Yaskawa INFORM job: -DEFRO-70-PRZYLACZE-70KASUJ.JBI

/JOB
//NAME -DEFRO-70-PRZYLACZE-70KASUJ
//POS
///NPOS 124,124,124,0,0,0
///TOOL 0
///POSTYPE PULSE
///PULSE
C00000=-283,-101162,-84213,3710,-80188,-1936
C00001=-283,-101162,-84213,3710,-80188,-1936
C00002=116617,-39062,-41553,1138,-40446,20
C00003=129312,23670,-33720,-14256,-61435,76595
C00004=149817,31841,-31795,27011,-57385,28137
C00005=152773,60456,-9717,30826,-76450,24874
C00006=149980,46799,-17890,30362,-63313,13597
C00007=141160,51169,-7378,14366,-65778,3091
C00008=136677,64016,6397,6150,-76179,-494
C00009=141378,9053,-49023,24268,-47565,-67133
C00010=125496,48327,-10508,-10752,-65084,-13725
C00011=130369,56785,-528,-1011,-71593,-13969
C00012=129107,53038,-4370,-2924,-69346,-18638
C00013=128986,13733,-25067,-13195,-71631,75488
C00014=115254,13128,-25616,-11802,-73565,79847
C00015=115259,22487,-34865,-12640,-63289,80918
C00016=131340,5225,-55572,19882,-37557,40272
C00017=141113,50251,-21422,35156,-71250,27064
C00018=141007,50182,-21498,35193,-71206,27085
C00019=141007,50182,-21498,35193,-71206,27085
C00020=137714,37646,-27763,32896,-58429,16473
C00021=129076,45247,-14016,15951,-62855,6645
C00022=121365,54735,-2868,3704,-70570,-4230
C00023=105889,56250,-7649,-21324,-75365,-25403
C00024=98023,31978,-40039,-45182,-56261,-13451
C00025=100224,44212,-25129,-32797,-73818,-42058
C00026=102299,40629,-26008,-28475,-71942,-45909
C00027=121076,21343,-35316,908,-62246,-81562
C00028=121076,10747,-22159,833,-75786,-81463
C00029=100383,18918,-18562,-9881,-76761,84439
C00030=101335,27463,-29788,-10664,-65529,85098
C00031=115713,4222,-56662,15198,-34727,46918
C00032=128373,44829,-27529,39504,-66240,29595
C00033=124328,33310,-32072,34883,-53820,19937
C00034=124328,33310,-32072,34883,-53820,19937
C00035=116075,45486,-13239,16661,-61560,10020
C00036=112317,60890,2820,11495,-73723,-606
C00037=94613,64601,2142,-17801,-79259,-22601
C00038=91137,54103,-11116,-25365,-70739,-18946
C00039=86945,42270,-27280,-36642,-61219,-13206
C00040=88301,54680,-13566,-28329,-78742,-39649
C00041=93612,48687,-14019,-16896,-75888,-44120
C00042=107037,24185,-32573,2312,-62235,-77114
C00043=100383,18918,-18562,-9881,-76761,84439
C00044=88082,30336,-7531,-8088,-78954,88284
C00045=89154,35127,-22112,-8522,-65087,85240
C00046=89544,34712,-22538,-8576,-65002,85121
C00047=100203,10236,-51959,9142,-32676,54086
C00048=115214,43849,-28542,43438,-61422,32379
C00049=110430,34623,-30597,35948,-49426,23884
C00050=101177,66932,10039,13677,-73518,2856
C00051=84754,73517,14044,-12253,-80824,-22539
C00052=78238,80066,13225,-23326,-87649,-28956
C00053=78238,80066,13225,-23326,-87649,-28956
C00054=77744,70007,4024,-24183,-84112,-37607
C00055=93905,32013,-24678,3546,-62668,-72921
C00056=93951,24843,-16667,3331,-71267,-72683
C00057=77831,45702,7684,-6459,-81284,91476
C00058=78073,52891,-3303,-6771,-70880,91958
C00059=86321,21390,-41402,2747,-32621,60915
C00060=102328,48592,-23384,46468,-56980,35399
C00061=97622,41313,-23800,35801,-45769,27976
C00062=95336,65754,6791,24352,-65412,15878
C00063=90551,78368,23842,15429,-74357,6364
C00064=75321,97136,42564,-11419,-90206,-17945
C00065=66680,76750,12803,-30175,-73528,-10031
C00066=68858,90162,29080,-20673,-90872,-36103
C00067=68858,90162,29080,-20673,-90872,-36103
C00068=68890,88039,27277,-20264,-89888,-36525
C00069=82457,45121,-10983,4500,-63864,-69204
C00070=77831,46763,5255,-6493,-79257,91580
C00071=100383,18918,-18562,-9881,-76761,84439
C00072=124101,-43184,-98243,-16518,52281,7000
C00073=123755,-7958,-89511,-14194,64535,5137
C00074=123755,-7958,-89511,-14194,64535,5137
C00075=120912,-12617,-93089,-9839,60859,10956
C00076=121533,-31212,-92910,-11510,35078,6544
C00077=122206,-29072,-90087,-12243,35589,-2657
C00078=123755,-7840,-89515,-14187,64596,5129
C00079=123755,-27930,-86554,-16069,52849,6788
C00080=123755,-31596,-85257,-16659,50271,7220
C00081=123755,-28371,-86416,-16134,52549,6837
C00082=123755,-7958,-89511,-14194,64535,5137
C00083=121932,-4467,-89644,-7852,68214,10996
C00084=130594,-5675,-87742,-32640,65606,16968
C00085=121207,-33956,-80021,-42944,8634,21416
C00086=121398,-33051,-89073,-12931,27077,-1891
C00087=119830,-29976,-89766,-6946,33011,-10480
C00088=121383,9671,-86957,-7975,82780,3273
C00089=123844,-33214,-84175,-16864,48398,7942
C00090=123999,-39711,-94755,-16482,51917,7023
C00091=123520,-8018,-89739,-13952,64610,5074
C00092=123514,-7754,-89533,-13967,64621,5071
C00093=125747,-8511,-91196,-20044,64124,16767
C00094=124758,-33497,-85798,-35788,21508,19109
C00095=121444,-34263,-87472,-15236,22128,1720
C00096=117635,-29901,-89670,2040,32900,-12364
C00097=120806,-19229,-91385,-7013,51591,-4269
C00098=123278,-3298,-89359,-12226,69976,6390
C00099=123735,-32674,-90978,-15994,53118,6740
C00100=123835,-44294,-91959,-17334,47983,7666
C00101=122869,-6543,-89983,-11258,66473,7782
C00102=122869,-6622,-89981,-11262,66432,7786
C00103=120666,-24161,-92251,-9656,44301,18332
C00104=120622,-35099,-88572,-13686,22135,5149
C00105=121670,-32826,-90694,-12460,29863,-58
C00106=120799,-29821,-90097,-9101,34108,-7769
C00107=117992,-25289,-89559,-1030,40191,-9143
C00108=122619,-6933,-90139,-10800,66466,8097
C00109=122622,-7156,-90314,-10803,66459,8098
C00110=123632,-25499,-87776,-15569,54758,6451
C00111=123637,-32760,-85682,-16630,49927,7238
C00112=123766,-34030,-92143,-16017,53144,6747
C00113=122032,-5500,-90078,-8484,67787,10331
C00114=122032,-5500,-90078,-8484,67787,10331
C00115=119888,-26436,-91823,-7086,40086,20761
C00116=120072,-35228,-83770,-17836,12895,7656
C00117=119245,-35145,-84473,-5873,14566,-1771
C00118=120774,-28613,-91055,-8481,37254,-8445
C00119=122137,-20625,-91389,-11840,49625,-8457
C00120=122281,3827,-88512,-9548,77692,7214
C00121=124756,-84422,-108366,-22045,38231,10349
C00122=2454,-100942,-83171,2490,-79441,1084
C00123=-283,-101162,-84213,3710,-80188,-1936
BC00000=570125
BC00001=954451
BC00002=878037
BC00003=914864
BC00004=914864
BC00005=914864
BC00006=914864
BC00007=914864
BC00008=914864
BC00009=914864
BC00010=914864
BC00011=914864
BC00012=914864
BC00013=914864
BC00014=914864
BC00015=914864
BC00016=914864
BC00017=914864
BC00018=914864
BC00019=914864
BC00020=914864
BC00021=914864
BC00022=914864
BC00023=914864
BC00024=914864
BC00025=914864
BC00026=914864
BC00027=914864
BC00028=914864
BC00029=914864
BC00030=914864
BC00031=914864
BC00032=914864
BC00033=914864
BC00034=914864
BC00035=914864
BC00036=914864
BC00037=914863
BC00038=914863
BC00039=914864
BC00040=914864
BC00041=914864
BC00042=914864
BC00043=914864
BC00044=914864
BC00045=914864
BC00046=914864
BC00047=914864
BC00048=914864
BC00049=914864
BC00050=914864
BC00051=914864
BC00052=914864
BC00053=914864
BC00054=914864
BC00055=914864
BC00056=914864
BC00057=914864
BC00058=914864
BC00059=914864
BC00060=914864
BC00061=914864
BC00062=914864
BC00063=914864
BC00064=914863
BC00065=914864
BC00066=914864
BC00067=914864
BC00068=914864
BC00069=914864
BC00070=914864
BC00071=914864
BC00072=869720
BC00073=869720
BC00074=869720
BC00075=869720
BC00076=869720
BC00077=869720
BC00078=869720
BC00079=869720
BC00080=869720
BC00081=908129
BC00082=908129
BC00083=908129
BC00084=907961
BC00085=908580
BC00086=908293
BC00087=908102
BC00088=907757
BC00089=908179
BC00090=945847
BC00091=945846
BC00092=945847
BC00093=946325
BC00094=946857
BC00095=946662
BC00096=946390
BC00097=946210
BC00098=945983
BC00099=945983
BC00100=984509
BC00101=984509
BC00102=984509
BC00103=984689
BC00104=985047
BC00105=984920
BC00106=984769
BC00107=984449
BC00108=984290
BC00109=984290
BC00110=984290
BC00111=1022837
BC00112=1022864
BC00113=1022864
BC00114=1022864
BC00115=1022915
BC00116=1023549
BC00117=1023332
BC00118=1022983
BC00119=1022931
BC00120=1022837
BC00121=1022837
BC00122=1040800
BC00123=570125
EC00000=1166,0
EC00001=1166,0
EC00002=-1743,0
EC00003=-1741,0
EC00004=-1741,0
EC00005=-1741,0
EC00006=-1740,0
EC00007=-1740,0
EC00008=-1740,0
EC00009=-1740,0
EC00010=-1740,0
EC00011=-1740,0
EC00012=-1740,0
EC00013=-1741,0
EC00014=-1741,0
EC00015=-1741,0
EC00016=-1741,0
EC00017=-1741,0
EC00018=-1741,0
EC00019=-1741,0
EC00020=-1740,0
EC00021=-1740,0
EC00022=-1740,0
EC00023=-1740,0
EC00024=-1740,0
EC00025=-1741,0
EC00026=-1741,0
EC00027=-1740,0
EC00028=-1740,0
EC00029=-1741,0
EC00030=-1741,0
EC00031=-1741,0
EC00032=-1741,0
EC00033=-1741,0
EC00034=-1741,0
EC00035=-1740,0
EC00036=-1740,0
EC00037=-1741,0
EC00038=-1741,0
EC00039=-1740,0
EC00040=-1741,0
EC00041=-1741,0
EC00042=-1740,0
EC00043=-1741,0
EC00044=-1741,0
EC00045=-1741,0
EC00046=-1741,0
EC00047=-1741,0
EC00048=-1741,0
EC00049=-1741,0
EC00050=-1740,0
EC00051=-1741,0
EC00052=-1741,0
EC00053=-1741,0
EC00054=-1741,0
EC00055=-1740,0
EC00056=-1740,0
EC00057=-1741,0
EC00058=-1741,0
EC00059=-1741,0
EC00060=-1741,0
EC00061=-1741,0
EC00062=-1740,0
EC00063=-1740,0
EC00064=-1741,0
EC00065=-1740,0
EC00066=-1741,0
EC00067=-1741,0
EC00068=-1741,0
EC00069=-1740,0
EC00070=-1741,0
EC00071=-1741,0
EC00072=-85617,0
EC00073=-85617,0
EC00074=-85617,0
EC00075=-85617,0
EC00076=-85617,0
EC00077=-85617,0
EC00078=-85617,0
EC00079=-85617,0
EC00080=-85617,0
EC00081=-85617,0
EC00082=-85617,0
EC00083=-85617,0
EC00084=-85617,0
EC00085=-85617,0
EC00086=-85617,0
EC00087=-85617,0
EC00088=-85617,0
EC00089=-85617,0
EC00090=-85617,0
EC00091=-85617,0
EC00092=-85617,0
EC00093=-85617,0
EC00094=-85617,0
EC00095=-85617,0
EC00096=-85617,0
EC00097=-85617,0
EC00098=-85617,0
EC00099=-85617,0
EC00100=-85617,0
EC00101=-85617,0
EC00102=-85617,0
EC00103=-85617,0
EC00104=-85617,0
EC00105=-85617,0
EC00106=-85617,0
EC00107=-85617,0
EC00108=-85617,0
EC00109=-85617,0
EC00110=-85617,0
EC00111=-85617,0
EC00112=-85617,0
EC00113=-85617,0
EC00114=-85617,0
EC00115=-85617,0
EC00116=-85617,0
EC00117=-85617,0
EC00118=-85617,0
EC00119=-85617,0
EC00120=-85617,0
EC00121=-85617,0
EC00122=946,0
EC00123=1166,0
//INST
///DATE 2025/05/08 13:43
///COMM OZZ
///ATTR SC,RW
///GROUP1 RB1,BS1
///GROUP2 ST1
NOP
MOVJ C00000 BC00000 VJ=70.00 DEC=20  +MOVJ EC00000 VJ=70.00
MOVJ C00001 BC00001 VJ=40.00 DEC=20  +MOVJ EC00001 VJ=40.00
MOVJ C00002 BC00002 VJ=70.00 DEC=20  +MOVJ EC00002 VJ=70.00
MOVJ C00003 BC00003 VJ=80.00 DEC=20  +MOVJ EC00003 VJ=80.00
MACRO1 MJ#(0) ARGF10
WVON WEV#(2)
ARCON
MOVL C00004 BC00004 V=5.0 DEC=20  +MOVJ EC00004 VJ=80.00
MOVC C00005 BC00005 V=5.0 DEC=20  +MOVJ EC00005 VJ=80.00
WVON WEV#(1)
MOVC C00006 BC00006 V=5.0 DEC=20  +MOVJ EC00006 VJ=80.00
MOVC C00007 BC00007 V=5.0 DEC=20  +MOVJ EC00007 VJ=80.00
MOVC C00008 BC00008 V=5.0 DEC=20  +MOVJ EC00008 VJ=80.00
MOVC C00009 BC00009 V=5.0 DEC=20  +MOVJ EC00009 VJ=80.00
MOVL C00010 BC00010 V=5.0 DEC=20  +MOVJ EC00010 VJ=80.00
MOVC C00011 BC00011 V=5.0 DEC=20  +MOVJ EC00011 VJ=80.00
MOVL C00012 BC00012 V=5.0 DEC=20  +MOVJ EC00012 VJ=80.00
WVOF
ARCOF
MOVJ C00013 BC00013 VJ=80.00 DEC=20  +MOVJ EC00013 VJ=80.00
MOVJ C00014 BC00014 VJ=80.00 DEC=20  +MOVJ EC00014 VJ=80.00
MOVJ C00015 BC00015 VJ=80.00 DEC=20  +MOVJ EC00015 VJ=0.78
MACRO1 MJ#(0) ARGF10
WVON WEV#(2)
ARCON
MOVC C00016 BC00016 V=5.0 DEC=20  +MOVJ EC00016 VJ=40.00
MOVL C00017 BC00017 V=5.0 DEC=20  +MOVJ EC00017 VJ=40.00
WVON WEV#(1)
MOVC C00018 BC00018 V=1500.0 DEC=20  +MOVJ EC00018 VJ=40.00
MOVC C00019 BC00019 V=600.0 DEC=20  +MOVJ EC00019 VJ=40.00
MOVC C00020 BC00020 V=5.0 DEC=20  +MOVJ EC00020 VJ=40.00
MOVC C00021 BC00021 V=5.0 DEC=20  +MOVJ EC00021 VJ=100.00
MOVC C00022 BC00022 V=5.0 DEC=20  +MOVJ EC00022 VJ=40.00
MOVC C00023 BC00023 V=5.0 DEC=20  +MOVJ EC00023 VJ=40.00
MOVL C00024 BC00024 V=5.0 DEC=20  +MOVJ EC00024 VJ=40.00
WVON WEV#(2)
MOVC C00025 BC00025 V=5.0 DEC=20  +MOVJ EC00025 VJ=40.00
MOVC C00026 BC00026 V=5.0 DEC=20  +MOVJ EC00026 VJ=80.00
MOVC C00027 BC00027 V=5.0 DEC=20  +MOVJ EC00027 VJ=40.00
WVOF
ARCOF
MOVJ C00028 BC00028 VJ=80.00 DEC=20  +MOVJ EC00028 VJ=80.00
MOVJ C00029 BC00029 VJ=80.00 DEC=20  +MOVJ EC00029 VJ=80.00
MOVJ C00030 BC00030 VJ=80.00 DEC=20  +MOVJ EC00030 VJ=80.00
MACRO1 MJ#(0) ARGF10
WVON WEV#(2)
ARCON
MOVC C00031 BC00031 V=5.0 DEC=20  +MOVJ EC00031 VJ=80.00
MOVL C00032 BC00032 V=5.0 DEC=20  +MOVJ EC00032 VJ=80.00
WVON WEV#(1)
MOVC C00033 BC00033 V=5.0 DEC=20  +MOVJ EC00033 VJ=80.00
MOVL C00034 BC00034 V=5.0 DEC=20  +MOVJ EC00034 VJ=80.00
MOVC C00035 BC00035 V=5.0 DEC=20  +MOVJ EC00035 VJ=80.00
MOVC C00036 BC00036 V=5.0 DEC=20  +MOVJ EC00036 VJ=80.00
MOVC C00037 BC00037 V=5.0 DEC=20  +MOVJ EC00037 VJ=80.00
MOVC C00038 BC00038 V=5.0 DEC=20  +MOVJ EC00038 VJ=80.00
MOVL C00039 BC00039 V=5.0 DEC=20  +MOVJ EC00039 VJ=80.00
MOVC C00040 BC00040 V=5.0 DEC=20  +MOVJ EC00040 VJ=80.00
MOVC C00041 BC00041 V=5.0 DEC=20  +MOVJ EC00041 VJ=80.00
MOVC C00042 BC00042 V=5.0 DEC=20  +MOVJ EC00042 VJ=80.00
WVOF
ARCOF
MOVJ C00043 BC00043 VJ=80.00 DEC=20  +MOVJ EC00043 VJ=80.00
MOVJ C00044 BC00044 VJ=80.00 DEC=20  +MOVJ EC00044 VJ=80.00
MOVJ C00045 BC00045 VJ=80.00 DEC=20  +MOVJ EC00045 VJ=80.00
MOVC C00046 BC00046 V=5.0 DEC=20  +MOVJ EC00046 VJ=80.00
MACRO1 MJ#(0) ARGF10
WVON WEV#(2)
ARCON
MOVC C00047 BC00047 V=5.0 DEC=20  +MOVJ EC00047 VJ=80.00
MOVC C00048 BC00048 V=5.0 DEC=20  +MOVJ EC00048 VJ=80.00
WVON WEV#(1)
MOVC C00049 BC00049 V=5.0 DEC=20  +MOVJ EC00049 VJ=80.00
MOVC C00050 BC00050 V=5.0 DEC=20  +MOVJ EC00050 VJ=80.00
MOVC C00051 BC00051 V=5.0 DEC=20  +MOVJ EC00051 VJ=80.00
MOVL C00052 BC00052 V=5.0 DEC=20  +MOVJ EC00052 VJ=80.00
MOVC C00053 BC00053 V=5.0 DEC=20  +MOVJ EC00053 VJ=80.00
MOVC C00054 BC00054 V=5.0 DEC=20  +MOVJ EC00054 VJ=80.00
MOVC C00055 BC00055 V=5.0 DEC=20  +MOVJ EC00055 VJ=80.00
WVOF
ARCOF
MOVJ C00056 BC00056 VJ=80.00 DEC=20  +MOVJ EC00056 VJ=80.00
MOVJ C00057 BC00057 VJ=80.00 DEC=20  +MOVJ EC00057 VJ=80.00
MOVJ C00058 BC00058 VJ=80.00 DEC=20  +MOVJ EC00058 VJ=80.00
MACRO1 MJ#(0) ARGF10
WVON WEV#(2)
ARCON
MOVC C00059 BC00059 V=5.0 DEC=20  +MOVJ EC00059 VJ=80.00
MOVC C00060 BC00060 V=5.0 DEC=20  +MOVJ EC00060 VJ=80.00
WVON WEV#(1)
MOVC C00061 BC00061 V=5.0 DEC=20  +MOVJ EC00061 VJ=80.00
MOVC C00062 BC00062 V=5.0 DEC=20  +MOVJ EC00062 VJ=80.00
MOVC C00063 BC00063 V=5.0 DEC=20  +MOVJ EC00063 VJ=80.00
MOVC C00064 BC00064 V=5.0 DEC=20  +MOVJ EC00064 VJ=80.00
MOVL C00065 BC00065 V=5.0 DEC=20  +MOVJ EC00065 VJ=80.00
MOVC C00066 BC00066 V=5.0 DEC=20  +MOVJ EC00066 VJ=80.00
MOVC C00067 BC00067 V=5.0 DEC=20  +MOVJ EC00067 VJ=80.00
MOVC C00068 BC00068 V=5.0 DEC=20  +MOVJ EC00068 VJ=80.00
MOVC C00069 BC00069 V=5.0 DEC=20  +MOVJ EC00069 VJ=80.00
ARCOF
WVOF
MOVJ C00070 BC00070 VJ=80.00 DEC=20  +MOVJ EC00070 VJ=80.00
MOVJ C00071 BC00071 VJ=80.00 DEC=20  +MOVJ EC00071 VJ=80.00
MOVJ C00072 BC00072 VJ=40.00 DEC=20  +MOVJ EC00072 VJ=40.00
MOVJ C00073 BC00073 VJ=80.00 DEC=20  +MOVJ EC00073 VJ=80.00
MACRO1 MJ#(0) ARGF4
ARCON
MOVC C00074 BC00074 V=5.0 DEC=20  +MOVJ EC00074 VJ=80.00
MOVC C00075 BC00075 V=5.0 DEC=20  +MOVJ EC00075 VJ=80.00
MOVC C00076 BC00076 V=5.0 DEC=20  +MOVJ EC00076 VJ=80.00
MOVC C00077 BC00077 V=5.0 DEC=20  +MOVJ EC00077 VJ=80.00
MOVC C00078 BC00078 V=5.0 DEC=20  +MOVJ EC00078 VJ=80.00
ARCOF
MOVJ C00079 BC00079 VJ=80.00 DEC=20  +MOVJ EC00079 VJ=80.00
MOVJ C00080 BC00080 VJ=80.00 DEC=20  +MOVJ EC00080 VJ=80.00
MOVJ C00081 BC00081 VJ=80.00 DEC=20  +MOVJ EC00081 VJ=80.00
MOVJ C00082 BC00082 VJ=80.00 DEC=20  +MOVJ EC00082 VJ=80.00
MACRO1 MJ#(0) ARGF4
ARCON
MOVC C00083 BC00083 V=5.0 DEC=20  +MOVJ EC00083 VJ=80.00
MOVC C00084 BC00084 V=5.0 DEC=20  +MOVJ EC00084 VJ=80.00
MOVC C00085 BC00085 V=5.0 DEC=20  +MOVJ EC00085 VJ=80.00
MOVC C00086 BC00086 V=5.0 DEC=20  +MOVJ EC00086 VJ=80.00
MOVC C00087 BC00087 V=5.0 DEC=20  +MOVJ EC00087 VJ=80.00
MOVC C00088 BC00088 V=5.0 DEC=20  +MOVJ EC00088 VJ=80.00
ARCOF
MOVJ C00089 BC00089 VJ=80.00 DEC=20  +MOVJ EC00089 VJ=80.00
MOVJ C00090 BC00090 VJ=80.00 DEC=20  +MOVJ EC00090 VJ=80.00
MOVJ C00091 BC00091 VJ=80.00 DEC=20  +MOVJ EC00091 VJ=80.00
ARCON
MOVC C00092 BC00092 V=5.0 DEC=20  +MOVJ EC00092 VJ=80.00
MOVC C00093 BC00093 V=5.0 DEC=20  +MOVJ EC00093 VJ=80.00
MOVC C00094 BC00094 V=5.0 DEC=20  +MOVJ EC00094 VJ=80.00
MOVC C00095 BC00095 V=5.0 DEC=20  +MOVJ EC00095 VJ=80.00
MOVC C00096 BC00096 V=5.0 DEC=20  +MOVJ EC00096 VJ=80.00
MOVC C00097 BC00097 V=5.0 DEC=20  +MOVJ EC00097 VJ=80.00
MOVC C00098 BC00098 V=3.3 DEC=20  +MOVJ EC00098 VJ=80.00
ARCOF
MOVJ C00099 BC00099 VJ=80.00 DEC=20  +MOVJ EC00099 VJ=80.00
MOVJ C00100 BC00100 VJ=80.00 DEC=20  +MOVJ EC00100 VJ=80.00
MOVJ C00101 BC00101 VJ=80.00 DEC=20  +MOVJ EC00101 VJ=80.00
ARCON
MOVC C00102 BC00102 V=5.0 DEC=20  +MOVJ EC00102 VJ=80.00
MOVC C00103 BC00103 V=5.0 DEC=20  +MOVJ EC00103 VJ=80.00
MOVC C00104 BC00104 V=5.0 DEC=20  +MOVJ EC00104 VJ=80.00
MOVC C00105 BC00105 V=5.0 DEC=20  +MOVJ EC00105 VJ=80.00
MOVC C00106 BC00106 V=5.0 DEC=20  +MOVJ EC00106 VJ=80.00
MOVC C00107 BC00107 V=5.0 DEC=20  +MOVJ EC00107 VJ=80.00
MOVC C00108 BC00108 V=3.3 DEC=20  +MOVJ EC00108 VJ=80.00
MOVL C00109 BC00109 V=3.3 DEC=20  +MOVJ EC00109 VJ=80.00
ARCOF
MOVJ C00110 BC00110 VJ=80.00 DEC=20  +MOVJ EC00110 VJ=80.00
MOVJ C00111 BC00111 VJ=80.00 DEC=20  +MOVJ EC00111 VJ=80.00
MOVJ C00112 BC00112 VJ=80.00 DEC=20  +MOVJ EC00112 VJ=80.00
MOVJ C00113 BC00113 VJ=80.00 DEC=20  +MOVJ EC00113 VJ=80.00
TIMER T=0.20
ARCON
MOVC C00114 BC00114 V=5.0 DEC=20  +MOVJ EC00114 VJ=80.00
MOVC C00115 BC00115 V=5.0 DEC=20  +MOVJ EC00115 VJ=80.00
MOVC C00116 BC00116 V=5.0 DEC=20  +MOVJ EC00116 VJ=80.00
MOVC C00117 BC00117 V=5.0 DEC=20  +MOVJ EC00117 VJ=80.00
MOVC C00118 BC00118 V=5.0 DEC=20  +MOVJ EC00118 VJ=80.00
MOVC C00119 BC00119 V=5.0 DEC=20  +MOVJ EC00119 VJ=80.00
MOVC C00120 BC00120 V=5.0 DEC=20  +MOVJ EC00120 VJ=80.00
ARCOF
MOVJ C00121 BC00121 VJ=80.00 DEC=20  +MOVJ EC00121 VJ=80.00
MOVJ C00122 BC00122 VJ=40.00 DEC=20  +MOVJ EC00122 VJ=40.00
MOVJ C00123 BC00123 VJ=40.00 DEC=20  +MOVJ EC00123 VJ=40.00
END
